Universal Robots URScript: T014_mistralai_Devstral-Small-2-24B-Instruct-2512_baseline_rep1_retry2.urscript

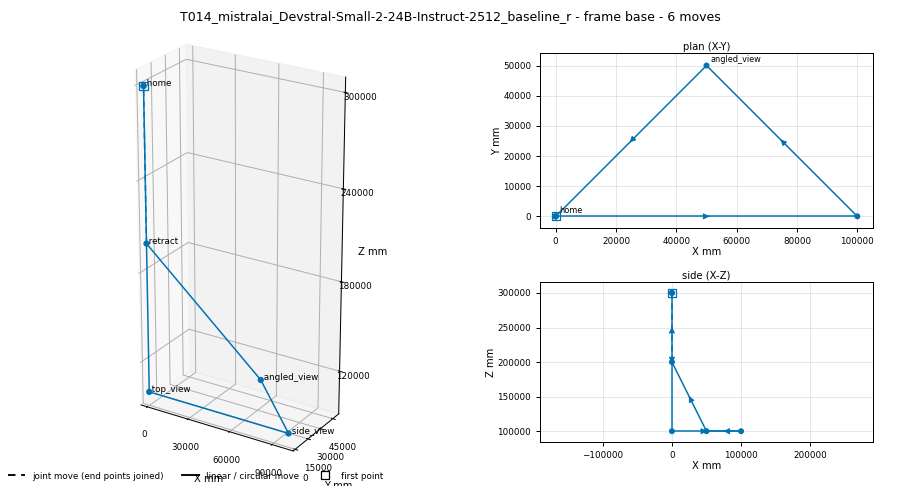
[picture p0: tool path of T014_mistralai_Devstral-Small-2-24B-Instruct-2512_baseline_rep1_retry2.urscript in frame base, 6 of 6 moves have a stored position in this frame; points joined in program order, loops and branches not executed]
def hybrid_inspection():
    # Define tool and base frames
    tool0 = p[0, 0, 0, 0, 0, 0]
    base = p[0, 0, 0, 0, 0, 0]

    # Define waypoints
    home = p[0, 0, 300, 0, 0, 0]
    top_view = p[0, 0, 100, 0, 0, 0]
    side_view = p[100, 0, 100, 0, 0, 0]
    angled_view = p[50, 50, 100, 0, 0, 0]
    retract = p[0, 0, 200, 0, 0, 0]

    # Set payload
    set_payload(0.4, p[0, 0, 0.1])

    # Move to home position
    movej(home, a=1.57, v=180.0, t=0, r=0)

    # Top-down view
    movel(top_view, a=1.57, v=150.0, t=0, r=0)

    # Side view
    movel(side_view, a=1.57, v=120.0, t=0, r=0)

    # Angled view
    movel(angled_view, a=1.57, v=120.0, t=0, r=0)

    # Retract
    movel(retract, a=1.57, v=180.0, t=0, r=0)

    # Return to home
    movej(home, a=1.57, v=180.0, t=0, r=0)

hybrid_inspection()
